# B&R Automation Studio project DriveControl
Automation Studio 4.5.2.102; Default project; technology packages: Acp10Arnc0 5.2.1

## Configuration SampleText

CPU 4PP065.0571-P74, AutomationRuntime D4.52, Build 4.1.2, Vc V4.25.0, Safety 1.6

### Task classes (Cpu.sw)
```
Cyclic#4:
  Program <- Program.prg
Libraries: sys_lib, Runtime, asstring, brsystem, AsBrStr, Library
```

### Hardware
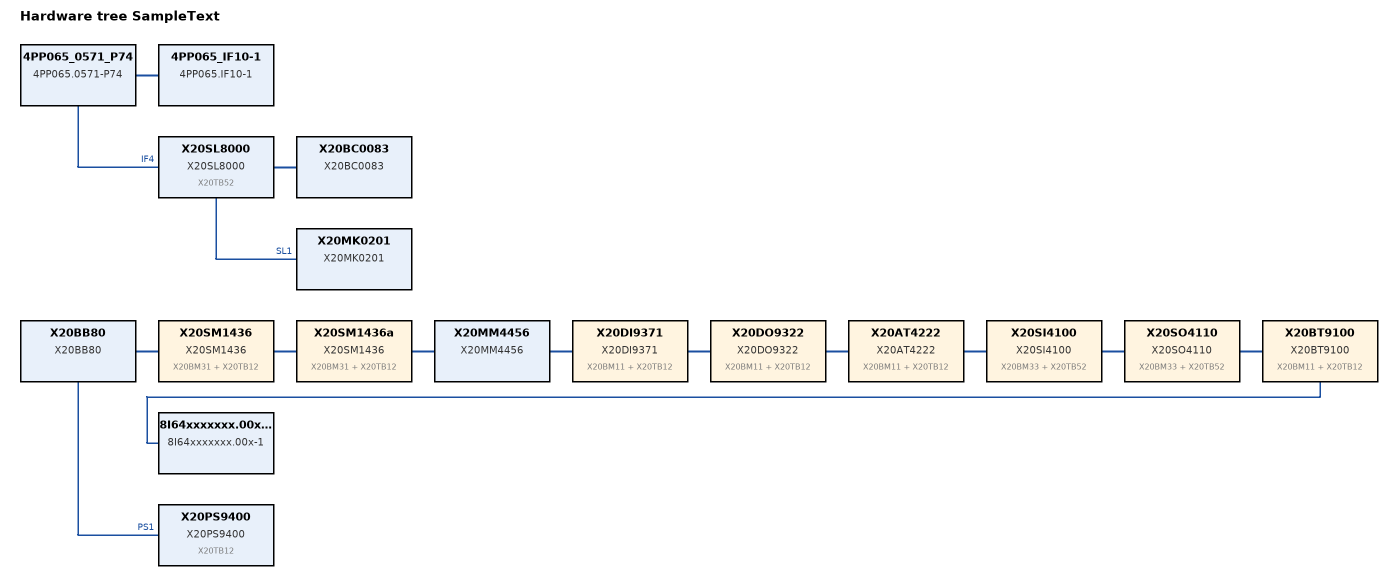
```
4PP065_0571_P74 : 4PP065.0571-P74 v1.1.2.0
  Connector IF5:
    ActivateDevice = 1
    Mode = Manual
    InternetAddress = 10.0.1.10
    SubnetMask = 255.255.255.0
  ConfigurationID = labBR
  TimerDeviceType = EPLX2X
  TimerDevice = 4PP065_0571_P74.IF4
  TaskClassIdleTime = 2000
  Cyclic1Duration = 2000
  Cyclic1Output = 1
4PP065_IF10-1 : 4PP065.IF10-1 v1.0.3.0  [SS -> 4PP065_0571_P74.SS1]
8I64xxxxxxx.00x-1 : 8I64xxxxxxx.00x-1 v1.3.9.1  [X2X1 -> X20BT9100.X2X1 [Cable Type=X2XCable, Length=10, Version=1.0.0.2]]
  packedETAD = packed
  packedETI = packed
  packedCMDD = packed
  packedCMI = packed
  ACC = 30
  DEC = 30
  UNS = 220
  NCR = 10
  NSP = 890
  COS = 64
  RSC = 33000
X20AT4222 : X20AT4222 v1.2.3.0  [SS1 -> X20TB12e.SS; SL -> X20BM11c.SL1]
X20BB80 : X20BB80 v1.0.2.0
X20BC0083 : X20BC0083 v2.9.0.0  [PLK1 -> X20SL8000.PLK2 (NodeNumber=2) [Cable Type=PowerlinkCable, Length=10, Version=1.0.0.2]; SL -> X20BB80.SL1]
X20BM11 : X20BM11 v1.0.0.1  [X2X1 -> X20BM33a.X2X2]
X20BM11a : X20BM11 v1.0.0.1  [X2X1 -> X20MM4456.X2X2]
X20BM11b : X20BM11 v1.0.0.1  [X2X1 -> X20BM11a.X2X2]
X20BM11c : X20BM11 v1.0.0.1  [X2X1 -> X20BM11b.X2X2]
X20BM31 : X20BM31 v1.0.0.1  [X2X1 -> X20BB80.IF1]
X20BM31a : X20BM31 v1.0.0.1  [X2X1 -> X20BM31.X2X2]
X20BM33 : X20BM33 v1.0.0.4  [X2X1 -> X20BM11c.X2X2]
X20BM33a : X20BM33 v1.0.0.4  [X2X1 -> X20BM33.X2X2]
X20BT9100 : X20BT9100 v1.0.3.0  [SS1 -> X20TB12f.SS; SL -> X20BM11.SL1]
X20DI9371 : X20DI9371 v1.0.2.0  [SS1 -> X20TB12c.SS; SL -> X20BM11a.SL1]
X20DO9322 : X20DO9322 v1.0.3.0  [SS1 -> X20TB12d.SS; SL -> X20BM11b.SL1]
X20MK0201 : X20MK0201 v1.0.0.0  [SL -> X20SL8000.SL1]
X20MM4456 : X20MM4456 v1.1.5.0  [X2X1 -> X20BM31a.X2X2]
X20PS9400 : X20PS9400 v1.0.2.4  [SS1 -> X20TB12.SS; PS -> X20BB80.PS1]
X20SI4100 : X20SI4100 v1.10.1.1  [SS1 -> X20TB52.SS; SL -> X20BM33.SL1]
X20SL8000 : X20SL8000 v1.6.5.1  [PLK1 -> 4PP065_0571_P74.IF4 (NodeNumber=1) [Cable Type=PowerlinkCable, Length=10, Version=1.0.0.2]; PLK2 -> X20BC0083.PLK1 (NodeNumber=1) [Cable Type=PowerlinkCable, Length=10, Version=1.0.0.2]; SS1 -> X20TB52b.SS]
  SafeProject = SafeLOGIC-1
X20SM1436 : X20SM1436 v2.3.0.0  [SS1 -> X20TB12a.SS; SL -> X20BM31.SL1]
X20SM1436a : X20SM1436 v2.3.0.0  [SS1 -> X20TB12b.SS; SL -> X20BM31a.SL1]
X20SO4110 : X20SO4110 v1.10.1.1  [SS1 -> X20TB52a.SS; SL -> X20BM33a.SL1]
  SafeModuleID = 3
X20TB12 : X20TB12 v1.0.0.0
X20TB12a : X20TB12 v1.0.0.0
X20TB12b : X20TB12 v1.0.0.0
X20TB12c : X20TB12 v1.0.0.0
X20TB12d : X20TB12 v1.0.0.0
X20TB12e : X20TB12 v1.0.0.0
X20TB12f : X20TB12 v1.0.0.0
X20TB52 : X20TB52 v1.0.0.1
X20TB52a : X20TB52 v1.0.0.1
X20TB52b : X20TB52 v1.0.0.1
```

### IoMap.iom - 4PP065_0571_P74/IoMap.iom
```iecst
VAR_CONFIG
	::stateMachine.speed AT %QW."8I64xxxxxxx.00x-1".LFRD_Output;
	::stateMachine.state AT %IW."8I64xxxxxxx.00x-1".ETAD_Input;
	::stateMachine.command AT %QW."8I64xxxxxxx.00x-1".CMDD_Output;
	::doorSM.direction AT %IX."X20DI9371".DigitalInput01;
	::doorSM.sw1 AT %IX."X20DI9371".DigitalInput02;
	::doorSM.sw2 AT %IX."X20DI9371".DigitalInput03;
	::doorSM.sw3 AT %IX."X20DI9371".DigitalInput04;
	::doorSM.sw4 AT %IX."X20DI9371".DigitalInput05;
	::ledSM.led1 AT %QX."X20DO9322".DigitalOutput02;
	::ledSM.led2 AT %QX."X20DO9322".DigitalOutput03;
	::ledSM.led3 AT %QX."X20DO9322".DigitalOutput04;
	::ledSM.led4 AT %QX."X20DO9322".DigitalOutput05;
END_VAR
```

- Physical/SampleText/4PP065_0571_P74/PvMap.vvm: same as Physical/SampleText/4PP065_0571_P74/Cpu.per
## Configuration Simulation

CPU , AutomationRuntime J4.25

### Task classes (Cpu.sw)
```
Libraries: AsIecCon, astime
```

### Hardware
```
PC_any : PC_any v1.1.0.0 (OrderNumber=PC)
```

- Physical/Simulation/PC_any/Cpu.per: same as Physical/SampleText/4PP065_0571_P74/Cpu.per
- Physical/Simulation/PC_any/PvMap.vvm: same as Physical/Simulation/PC_any/IOMap.iom
## Logical view

Binary libraries used (declarations not repeated): RUNTIME, OPERATOR, AsIecCon, astime, sys_lib, asstring, brsystem, AsBrStr

### Global.var - Global variables
```iecst
VAR
	doorSM : DoorStateMashine := (0);
	ledSM : LedStateMashine := (0);
	stateMachine : DriveStateMashine := (0);
END_VAR
```


### Library Logical/Library (ANSIC)

#### Types.typ - Exported data types
```iecst
TYPE
	DoorStates :
		(
		ST_INIT,
		ST_UNKNOWN,
		ST_OPEN,
		ST_CLOSE,
		ST_ACC_POS,
		ST_ACC_NEG,
		ST_POS,
		ST_NEG,
		ST_DEC_POS,
		ST_DEC_NEG
		);
END_TYPE
```

#### Constants.var - Exported constants
```iecst
VAR CONSTANT
	SPEED_SLOW : INT := 300; (*Slow speed: S0-S1, S2-S3, position search*)
	SPEED_FAST : INT := 800; (*Fast speed: S1-S2*)
	SPEED_STOP : INT := 0;
	DRV_STATE_MASK : UINT := 16#006F; (*Status word mask*)
	STATE_SWITCHED_ON : UINT := 16#0021; (*Ready to switch on*)
	STATE_READY : UINT := 16#0023; (*Switched on*)
	STATE_ENABLED : UINT := 16#0027; (*Operation enabled*)
	STATE_FAULT_BIT : UINT := 16#0008; (*Fault bit*)
	CMD_SHUTDOWN : UINT := 16#0006;
	CMD_SWITCH_ON : UINT := 16#0007;
	CMD_ENABLE : UINT := 16#000F;
	CMD_FAULT_RESET : UINT := 16#0080;
	BLINK_HALF_PERIOD_MS : UDINT := 500; (*1 Hz blink*)
END_VAR
```

#### Library.fun - Exported functions and function blocks
```iecst
{REDUND_ERROR} FUNCTION_BLOCK DriveStateMashine (*Frequency inverter control (CiA402)*) (*$GROUP=User,$CAT=User,$GROUPICON=User.png,$CATICON=User.png*)
	VAR_INPUT
		state : UINT; (*Inverter status word (ETAD)*)
		enable : BOOL; (*Enable FB*)
		speedSet : INT; (*Speed setpoint from door logic*)
	END_VAR
	VAR_OUTPUT
		command : UINT; (*Inverter control word (CMDD)*)
		speed : INT; (*Speed to inverter (LFRD)*)
	END_VAR
END_FUNCTION_BLOCK

{REDUND_ERROR} FUNCTION_BLOCK DoorStateMashine (*Door state machine*) (*$GROUP=User,$CAT=User,$GROUPICON=User.png,$CATICON=User.png*)
	VAR_INPUT
		state : UINT; (*Inverter status word*)
		sw1 : BOOL; (*S0 - door open*)
		sw2 : BOOL; (*S1*)
		sw3 : BOOL; (*S2*)
		sw4 : BOOL; (*S3 - door closed*)
		direction : BOOL; (*Switch: 1 - close, 0 - open*)
	END_VAR
	VAR_OUTPUT
		speed : INT; (*Speed setpoint*)
		doorState : DoorStates; (*Current door state*)
	END_VAR
	VAR
		s0Prev : BOOL; (*Sensor levels on previous cycle*)
		s1Prev : BOOL;
		s2Prev : BOOL;
		s3Prev : BOOL;
	END_VAR
END_FUNCTION_BLOCK

{REDUND_ERROR} FUNCTION_BLOCK LedStateMashine (*LED indication*) (*$GROUP=User,$CAT=User,$GROUPICON=User.png,$CATICON=User.png*)
	VAR_INPUT
		state : UINT; (*Door state*)
		cycleTime : UDINT; (*Task cycle time, ms*)
	END_VAR
	VAR_OUTPUT
		led1 : BOOL; (*S0*)
		led2 : BOOL; (*S1*)
		led3 : BOOL; (*S2*)
		led4 : BOOL; (*S3*)
		timer : INT; (*Blink timer, ms*)
	END_VAR
	VAR
		elapsed : UDINT;
		blink : BOOL;
	END_VAR
END_FUNCTION_BLOCK
```

#### DriveStateMashine.c
```c
#include <bur/plctypes.h>
#ifdef __cplusplus
	extern "C"
	{
#endif
#include "Library.h"
#ifdef __cplusplus
	};
#endif

void DriveStateMashine(struct DriveStateMashine* inst)
{
	UINT st = inst->state & DRV_STATE_MASK;

	if (!inst->enable)
	{
		inst->command = CMD_SHUTDOWN;
		inst->speed   = 0;
		return;
	}

	if (inst->state & STATE_FAULT_BIT)
	{
		inst->command = CMD_FAULT_RESET;
		inst->speed   = 0;
		return;
	}

	if (st == STATE_ENABLED)
	{
		inst->command = CMD_ENABLE;
		inst->speed   = inst->speedSet;
	}
	else if (st == STATE_READY)
	{
		inst->command = CMD_ENABLE;
		inst->speed   = 0;
	}
	else if (st == STATE_SWITCHED_ON)
	{
		inst->command = CMD_SWITCH_ON;
		inst->speed   = 0;
	}
	else
	{
		inst->command = CMD_SHUTDOWN;
		inst->speed   = 0;
	}
}
```

#### DoorStateMashine.c
```c
#include <bur/plctypes.h>
#ifdef __cplusplus
	extern "C"
	{
#endif
	#include "Library.h"
#ifdef __cplusplus
	};
#endif

void DoorStateMashine(struct DoorStateMashine* inst)
{
	BOOL s0 = inst->sw1;
	BOOL s1 = inst->sw2;
	BOOL s2 = inst->sw3;
	BOOL s3 = inst->sw4;

	BOOL s0Changed = (s0 != inst->s0Prev);
	BOOL s1Changed = (s1 != inst->s1Prev);
	BOOL s2Changed = (s2 != inst->s2Prev);
	BOOL s3Changed = (s3 != inst->s3Prev);

	BOOL driveOn = ((inst->state & DRV_STATE_MASK) == STATE_ENABLED);
	DoorStates stateAtStart;

	if (!driveOn && inst->doorState != ST_INIT)
		inst->doorState = ST_INIT;

	stateAtStart = inst->doorState;

	switch (inst->doorState)
	{
		case ST_INIT:
			inst->speed = SPEED_STOP;
			if (driveOn)
				inst->doorState = ST_UNKNOWN;
			break;

		case ST_UNKNOWN:
			inst->speed = inst->direction ? SPEED_SLOW : -SPEED_SLOW;
			if (!inst->direction && s0Changed)
				inst->doorState = ST_OPEN;
			else if (inst->direction && s3Changed)
				inst->doorState = ST_CLOSE;
			break;

		case ST_OPEN:
			inst->speed = SPEED_STOP;
			if (inst->direction)
				inst->doorState = ST_ACC_POS;
			break;

		case ST_ACC_POS:
			inst->speed = SPEED_SLOW;
			if (!inst->direction)
				inst->doorState = ST_DEC_NEG;
			else if (s1Changed)
				inst->doorState = ST_POS;
			break;

		case ST_POS:
			inst->speed = SPEED_FAST;
			if (!inst->direction)
				inst->doorState = ST_NEG;
			else if (s2Changed)
				inst->doorState = ST_DEC_POS;
			break;

		case ST_DEC_POS:
			inst->speed = SPEED_SLOW;
			if (!inst->direction)
				inst->doorState = ST_ACC_NEG;
			else if (s3Changed)
				inst->doorState = ST_CLOSE;
			break;

		case ST_CLOSE:
			inst->speed = SPEED_STOP;
			if (!inst->direction)
				inst->doorState = ST_ACC_NEG;
			break;

		case ST_ACC_NEG:
			inst->speed = -SPEED_SLOW;
			if (inst->direction)
				inst->doorState = ST_DEC_POS;
			else if (s2Changed)
				inst->doorState = ST_NEG;
			break;

		case ST_NEG:
			inst->speed = -SPEED_FAST;
			if (inst->direction)
				inst->doorState = ST_POS;
			else if (s1Changed)
				inst->doorState = ST_DEC_NEG;
			break;

		case ST_DEC_NEG:
			inst->speed = -SPEED_SLOW;
			if (inst->direction)
				inst->doorState = ST_ACC_POS;
			else if (s0Changed)
				inst->doorState = ST_OPEN;
			break;

		default:
			inst->speed = SPEED_STOP;
			inst->doorState = ST_INIT;
			break;
	}

	if (stateAtStart == ST_INIT || inst->doorState == ST_INIT)
	{
		inst->s0Prev = 0;
		inst->s1Prev = 0;
		inst->s2Prev = 0;
		inst->s3Prev = 0;
	}
	else
	{
		inst->s0Prev = s0;
		inst->s1Prev = s1;
		inst->s2Prev = s2;
		inst->s3Prev = s3;
	}
}
```

#### LedStateMashine.c
```c
#include <bur/plctypes.h>
#ifdef __cplusplus
	extern "C"
	{
#endif
	#include "Library.h"
#ifdef __cplusplus
	};
#endif

static void SetLeds(struct LedStateMashine* inst, BOOL l1, BOOL l2, BOOL l3, BOOL l4)
{
	inst->led1 = l1;
	inst->led2 = l2;
	inst->led3 = l3;
	inst->led4 = l4;
}

void LedStateMashine(struct LedStateMashine* inst)
{
	UDINT dt = inst->cycleTime;
	if (dt == 0)
		dt = 100;

	switch (inst->state)
	{
		case ST_UNKNOWN:
			inst->elapsed += dt;
			if (inst->elapsed >= BLINK_HALF_PERIOD_MS)
			{
				inst->elapsed = 0;
				inst->blink = !inst->blink;
			}
			SetLeds(inst, inst->blink, inst->blink, inst->blink, inst->blink);
			break;

		case ST_OPEN:     SetLeds(inst, 0, 0, 0, 0); break;
		case ST_ACC_POS:  SetLeds(inst, 1, 0, 0, 0); break;
		case ST_POS:      SetLeds(inst, 1, 1, 0, 0); break;
		case ST_DEC_POS:  SetLeds(inst, 1, 1, 1, 0); break;
		case ST_CLOSE:    SetLeds(inst, 1, 1, 1, 1); break;
		case ST_ACC_NEG:  SetLeds(inst, 1, 1, 1, 0); break;
		case ST_NEG:      SetLeds(inst, 1, 1, 0, 0); break;
		case ST_DEC_NEG:  SetLeds(inst, 1, 0, 0, 0); break;

		case ST_INIT:
		default:
			SetLeds(inst, 0, 0, 0, 0);
			break;
	}

	if (inst->state != ST_UNKNOWN)
	{
		inst->elapsed = 0;
		inst->blink = 0;
	}
	inst->timer = (INT)inst->elapsed;
}
```

### Program Logical/Program (ANSIC)

#### Main.c - Init, cyclic, exit code
```c
#include <bur/plctypes.h>

#ifdef _DEFAULT_INCLUDES
	#include <AsDefault.h>
#endif

static RTInfo_typ rtInfo;

void _INIT ProgramInit(void)
{
	rtInfo.enable = 1;
	RTInfo(&rtInfo);
	ledSM.cycleTime = rtInfo.cycle_time / 1000;
	if (ledSM.cycleTime == 0)
		ledSM.cycleTime = 100;

	stateMachine.enable   = 0;
	stateMachine.speedSet = 0;
	stateMachine.command  = CMD_SHUTDOWN;
	stateMachine.speed    = 0;

	doorSM.doorState = ST_INIT;
	doorSM.speed     = 0;

	ledSM.state = ST_INIT;
	ledSM.led1  = 0;
	ledSM.led2  = 0;
	ledSM.led3  = 0;
	ledSM.led4  = 0;
}

void _CYCLIC ProgramCyclic(void)
{
	doorSM.state = stateMachine.state;
	DoorStateMashine(&doorSM);

	stateMachine.enable   = 1;
	stateMachine.speedSet = doorSM.speed;
	DriveStateMashine(&stateMachine);

	ledSM.state = (UINT)doorSM.doorState;
	LedStateMashine(&ledSM);
}
```
